    IF ((x0 = FALSE) AND  (x1 = FALSE) AND  (x2 = FALSE) AND  (t0.Q = FALSE)) THEN 
        cstate58 := 7390; y0 := FALSE; y1 := TRUE; t0_start := FALSE; 
    ELSIF ((x0 = FALSE) AND  (x1 = FALSE) AND  (x2 = FALSE) AND  (t0.Q = TRUE)) THEN 
        cstate58 := 7378; y0 := FALSE; y1 := TRUE; t0_start := FALSE; 
    ELSIF ((x0 = FALSE) AND  (x1 = FALSE) AND  (x2 = TRUE) AND  (t0.Q = FALSE)) THEN 
        cstate58 := 7582; y0 := FALSE; y1 := TRUE; t0_start := FALSE; 
    ELSIF ((x0 = FALSE) AND  (x1 = FALSE) AND  (x2 = TRUE) AND  (t0.Q = TRUE)) THEN 
        cstate58 := 7570; y0 := FALSE; y1 := TRUE; t0_start := FALSE; 
    ELSIF ((x0 = FALSE) AND  (x1 = TRUE) AND  (x2 = FALSE) AND  (t0.Q = FALSE)) THEN 
        cstate58 := 6340; y0 := FALSE; y1 := FALSE; t0_start := FALSE; 
    ELSIF ((x0 = FALSE) AND  (x1 = TRUE) AND  (x2 = FALSE) AND  (t0.Q = TRUE)) THEN 
        cstate58 := 6338; y0 := FALSE; y1 := FALSE; t0_start := FALSE; 
    ELSIF ((x0 = FALSE) AND  (x1 = TRUE) AND  (x2 = TRUE) AND  (t0.Q = FALSE)) THEN 
        cstate58 := 6532; y0 := FALSE; y1 := FALSE; t0_start := FALSE; 
    ELSIF ((x0 = FALSE) AND  (x1 = TRUE) AND  (x2 = TRUE) AND  (t0.Q = TRUE)) THEN 
        cstate58 := 6530; y0 := FALSE; y1 := FALSE; t0_start := FALSE; 
    ELSIF ((x0 = TRUE) AND  (x1 = FALSE) AND  (x2 = FALSE) AND  (t0.Q = FALSE)) THEN 
        cstate58 := 5192; y0 := TRUE; y1 := FALSE; t0_start := FALSE; 
    ELSIF ((x0 = TRUE) AND  (x1 = FALSE) AND  (x2 = FALSE) AND  (t0.Q = TRUE)) THEN 
        cstate58 := 5186; y0 := TRUE; y1 := FALSE; t0_start := FALSE; 
    ELSIF ((x0 = TRUE) AND  (x1 = FALSE) AND  (x2 = TRUE) AND  (t0.Q = FALSE)) THEN 
        cstate58 := 3848; y0 := FALSE; y1 := FALSE; t0_start := FALSE; 
    ELSIF ((x0 = TRUE) AND  (x1 = FALSE) AND  (x2 = TRUE) AND  (t0.Q = TRUE)) THEN 
        cstate58 := 3842; y0 := FALSE; y1 := FALSE; t0_start := FALSE; 
    ELSIF ((x0 = TRUE) AND  (x1 = TRUE) AND  (x2 = FALSE) AND  (t0.Q = FALSE)) THEN 
        cstate58 := 4678; y0 := TRUE; y1 := FALSE; t0_start := FALSE; 
    ELSIF ((x0 = TRUE) AND  (x1 = TRUE) AND  (x2 = FALSE) AND  (t0.Q = TRUE)) THEN 
        cstate58 := 4674; y0 := TRUE; y1 := FALSE; t0_start := FALSE; 
    ELSIF ((x0 = TRUE) AND  (x1 = TRUE) AND  (x2 = TRUE) AND  (t0.Q = FALSE)) THEN 
        cstate58 := 2502; y0 := FALSE; y1 := FALSE; t0_start := FALSE; 
    ELSIF ((x0 = TRUE) AND  (x1 = TRUE) AND  (x2 = TRUE) AND  (t0.Q = TRUE)) THEN 
        cstate58 := 2498; y0 := FALSE; y1 := FALSE; t0_start := FALSE; 
    END_IF;
6338:
    IF ((x0 = FALSE) AND  (x1 = FALSE) AND  (x2 = FALSE) AND  (t0.Q = FALSE)) THEN 
        cstate58 := 6340; y0 := FALSE; y1 := FALSE; t0_start := FALSE; 
    ELSIF ((x0 = FALSE) AND  (x1 = FALSE) AND  (x2 = FALSE) AND  (t0.Q = TRUE)) THEN 
        cstate58 := 6338; y0 := FALSE; y1 := FALSE; t0_start := FALSE; 
    ELSIF ((x0 = FALSE) AND  (x1 = FALSE) AND  (x2 = TRUE) AND  (t0.Q = FALSE)) THEN 
        cstate58 := 6468; y0 := FALSE; y1 := FALSE; t0_start := TRUE; t0_up := FALSE; 
    ELSIF ((x0 = FALSE) AND  (x1 = FALSE) AND  (x2 = TRUE) AND  (t0.Q = TRUE)) THEN 
        cstate58 := 6466; y0 := FALSE; y1 := FALSE; t0_start := TRUE; t0_up := FALSE; 
    ELSIF ((x0 = FALSE) AND  (x1 = TRUE) AND  (x2 = FALSE) AND  (t0.Q = FALSE)) THEN 
        cstate58 := 6340; y0 := FALSE; y1 := FALSE; t0_start := FALSE; 
    ELSIF ((x0 = FALSE) AND  (x1 = TRUE) AND  (x2 = FALSE) AND  (t0.Q = TRUE)) THEN 
        cstate58 := 6338; y0 := FALSE; y1 := FALSE; t0_start := FALSE; 
    ELSIF ((x0 = FALSE) AND  (x1 = TRUE) AND  (x2 = TRUE) AND  (t0.Q = FALSE)) THEN 
        cstate58 := 6468; y0 := FALSE; y1 := FALSE; t0_start := TRUE; t0_up := FALSE; 
    ELSIF ((x0 = FALSE) AND  (x1 = TRUE) AND  (x2 = TRUE) AND  (t0.Q = TRUE)) THEN 
        cstate58 := 6466; y0 := FALSE; y1 := FALSE; t0_start := TRUE; t0_up := FALSE; 
    ELSIF ((x0 = TRUE) AND  (x1 = FALSE) AND  (x2 = FALSE) AND  (t0.Q = FALSE)) THEN 
        cstate58 := 4168; y0 := TRUE; y1 := FALSE; t0_start := FALSE; 
    ELSIF ((x0 = TRUE) AND  (x1 = FALSE) AND  (x2 = FALSE) AND  (t0.Q = TRUE)) THEN 
        cstate58 := 4162; y0 := TRUE; y1 := FALSE; t0_start := FALSE; 
    ELSIF ((x0 = TRUE) AND  (x1 = FALSE) AND  (x2 = TRUE) AND  (t0.Q = FALSE)) THEN 
        cstate58 := 2760; y0 := FALSE; y1 := FALSE; t0_start := TRUE; t0_up := FALSE; 
    ELSIF ((x0 = TRUE) AND  (x1 = FALSE) AND  (x2 = TRUE) AND  (t0.Q = TRUE)) THEN 
        cstate58 := 2754; y0 := FALSE; y1 := FALSE; t0_start := TRUE; t0_up := FALSE; 
    ELSIF ((x0 = TRUE) AND  (x1 = TRUE) AND  (x2 = FALSE) AND  (t0.Q = FALSE)) THEN 
        cstate58 := 4678; y0 := TRUE; y1 := FALSE; t0_start := FALSE; 
    ELSIF ((x0 = TRUE) AND  (x1 = TRUE) AND  (x2 = FALSE) AND  (t0.Q = TRUE)) THEN 
        cstate58 := 4674; y0 := TRUE; y1 := FALSE; t0_start := FALSE; 
    ELSIF ((x0 = TRUE) AND  (x1 = TRUE) AND  (x2 = TRUE) AND  (t0.Q = FALSE)) THEN 
        cstate58 := 2566; y0 := FALSE; y1 := FALSE; t0_start := TRUE; t0_up := FALSE; 
    ELSIF ((x0 = TRUE) AND  (x1 = TRUE) AND  (x2 = TRUE) AND  (t0.Q = TRUE)) THEN 
        cstate58 := 2562; y0 := FALSE; y1 := FALSE; t0_start := TRUE; t0_up := FALSE; 
    END_IF;
1226:
    IF ((x0 = FALSE) AND  (x1 = FALSE) AND  (x2 = FALSE) AND  (t0.Q = FALSE)) THEN 
        cstate58 := 1238; y0 := FALSE; y1 := TRUE; t0_start := FALSE; 
    ELSIF ((x0 = FALSE) AND  (x1 = FALSE) AND  (x2 = FALSE) AND  (t0.Q = TRUE)) THEN 
        cstate58 := 1226; y0 := FALSE; y1 := TRUE; t0_start := FALSE; 
    ELSIF ((x0 = FALSE) AND  (x1 = FALSE) AND  (x2 = TRUE) AND  (t0.Q = FALSE)) THEN 
        cstate58 := 1368; y0 := FALSE; y1 := TRUE; t0_start := TRUE; t0_up := FALSE; 
    ELSIF ((x0 = FALSE) AND  (x1 = FALSE) AND  (x2 = TRUE) AND  (t0.Q = TRUE)) THEN 
        cstate58 := 1356; y0 := FALSE; y1 := TRUE; t0_start := TRUE; t0_up := FALSE; 
    ELSIF ((x0 = FALSE) AND  (x1 = TRUE) AND  (x2 = FALSE) AND  (t0.Q = FALSE)) THEN 
        cstate58 := 1220; y0 := FALSE; y1 := FALSE; t0_start := FALSE; 
    ELSIF ((x0 = FALSE) AND  (x1 = TRUE) AND  (x2 = FALSE) AND  (t0.Q = TRUE)) THEN 
        cstate58 := 1218; y0 := FALSE; y1 := FALSE; t0_start := FALSE; 
    ELSIF ((x0 = FALSE) AND  (x1 = TRUE) AND  (x2 = TRUE) AND  (t0.Q = FALSE)) THEN 
        cstate58 := 1348; y0 := FALSE; y1 := FALSE; t0_start := TRUE; t0_up := FALSE; 
    ELSIF ((x0 = FALSE) AND  (x1 = TRUE) AND  (x2 = TRUE) AND  (t0.Q = TRUE)) THEN 
        cstate58 := 1346; y0 := FALSE; y1 := FALSE; t0_start := TRUE; t0_up := FALSE; 
    ELSIF ((x0 = TRUE) AND  (x1 = FALSE) AND  (x2 = FALSE) AND  (t0.Q = FALSE)) THEN 
        cstate58 := 5192; y0 := TRUE; y1 := FALSE; t0_start := FALSE; 
    ELSIF ((x0 = TRUE) AND  (x1 = FALSE) AND  (x2 = FALSE) AND  (t0.Q = TRUE)) THEN 
        cstate58 := 5186; y0 := TRUE; y1 := FALSE; t0_start := FALSE; 
    ELSIF ((x0 = TRUE) AND  (x1 = FALSE) AND  (x2 = TRUE) AND  (t0.Q = FALSE)) THEN 
        cstate58 := 3784; y0 := FALSE; y1 := FALSE; t0_start := TRUE; t0_up := FALSE; 
    ELSIF ((x0 = TRUE) AND  (x1 = FALSE) AND  (x2 = TRUE) AND  (t0.Q = TRUE)) THEN 
        cstate58 := 3778; y0 := FALSE; y1 := FALSE; t0_start := TRUE; t0_up := FALSE; 
    ELSIF ((x0 = TRUE) AND  (x1 = TRUE) AND  (x2 = FALSE) AND  (t0.Q = FALSE)) THEN 
        cstate58 := 4678; y0 := TRUE; y1 := FALSE; t0_start := FALSE; 
    ELSIF ((x0 = TRUE) AND  (x1 = TRUE) AND  (x2 = FALSE) AND  (t0.Q = TRUE)) THEN 
        cstate58 := 4674; y0 := TRUE; y1 := FALSE; t0_start := FALSE; 
    ELSIF ((x0 = TRUE) AND  (x1 = TRUE) AND  (x2 = TRUE) AND  (t0.Q = FALSE)) THEN 
        cstate58 := 2566; y0 := FALSE; y1 := FALSE; t0_start := TRUE; t0_up := FALSE; 
    ELSIF ((x0 = TRUE) AND  (x1 = TRUE) AND  (x2 = TRUE) AND  (t0.Q = TRUE)) THEN 
        cstate58 := 2562; y0 := FALSE; y1 := FALSE; t0_start := TRUE; t0_up := FALSE; 
    END_IF;
7370:
    IF ((x0 = FALSE) AND  (x1 = FALSE) AND  (x2 = FALSE) AND  (t0.Q = FALSE)) THEN 
        cstate58 := 7382; y0 := FALSE; y1 := TRUE; t0_start := FALSE; 
    ELSIF ((x0 = FALSE) AND  (x1 = FALSE) AND  (x2 = FALSE) AND  (t0.Q = TRUE)) THEN 
        cstate58 := 7370; y0 := FALSE; y1 := TRUE; t0_start := FALSE; 
    ELSIF ((x0 = FALSE) AND  (x1 = FALSE) AND  (x2 = TRUE) AND  (t0.Q = FALSE)) THEN 
        cstate58 := 7512; y0 := FALSE; y1 := TRUE; t0_start := TRUE; t0_up := FALSE; 
    ELSIF ((x0 = FALSE) AND  (x1 = FALSE) AND  (x2 = TRUE) AND  (t0.Q = TRUE)) THEN 
        cstate58 := 7500; y0 := FALSE; y1 := TRUE; t0_start := TRUE; t0_up := FALSE; 
    ELSIF ((x0 = FALSE) AND  (x1 = TRUE) AND  (x2 = FALSE) AND  (t0.Q = FALSE)) THEN 
        cstate58 := 6340; y0 := FALSE; y1 := FALSE; t0_start := FALSE; 
    ELSIF ((x0 = FALSE) AND  (x1 = TRUE) AND  (x2 = FALSE) AND  (t0.Q = TRUE)) THEN 
        cstate58 := 6338; y0 := FALSE; y1 := FALSE; t0_start := FALSE; 
    ELSIF ((x0 = FALSE) AND  (x1 = TRUE) AND  (x2 = TRUE) AND  (t0.Q = FALSE)) THEN 
        cstate58 := 6468; y0 := FALSE; y1 := FALSE; t0_start := TRUE; t0_up := FALSE; 
    ELSIF ((x0 = FALSE) AND  (x1 = TRUE) AND  (x2 = TRUE) AND  (t0.Q = TRUE)) THEN 
        cstate58 := 6466; y0 := FALSE; y1 := FALSE; t0_start := TRUE; t0_up := FALSE; 
    ELSIF ((x0 = TRUE) AND  (x1 = FALSE) AND  (x2 = FALSE) AND  (t0.Q = FALSE)) THEN 
        cstate58 := 5192; y0 := TRUE; y1 := FALSE; t0_start := FALSE; 
    ELSIF ((x0 = TRUE) AND  (x1 = FALSE) AND  (x2 = FALSE) AND  (t0.Q = TRUE)) THEN 
        cstate58 := 5186; y0 := TRUE; y1 := FALSE; t0_start := FALSE; 
    ELSIF ((x0 = TRUE) AND  (x1 = FALSE) AND  (x2 = TRUE) AND  (t0.Q = FALSE)) THEN 
        cstate58 := 3784; y0 := FALSE; y1 := FALSE; t0_start := TRUE; t0_up := FALSE; 
    ELSIF ((x0 = TRUE) AND  (x1 = FALSE) AND  (x2 = TRUE) AND  (t0.Q = TRUE)) THEN 
        cstate58 := 3778; y0 := FALSE; y1 := FALSE; t0_start := TRUE; t0_up := FALSE; 
    ELSIF ((x0 = TRUE) AND  (x1 = TRUE) AND  (x2 = FALSE) AND  (t0.Q = FALSE)) THEN 
        cstate58 := 4678; y0 := TRUE; y1 := FALSE; t0_start := FALSE; 
    ELSIF ((x0 = TRUE) AND  (x1 = TRUE) AND  (x2 = FALSE) AND  (t0.Q = TRUE)) THEN 
        cstate58 := 4674; y0 := TRUE; y1 := FALSE; t0_start := FALSE; 
    ELSIF ((x0 = TRUE) AND  (x1 = TRUE) AND  (x2 = TRUE) AND  (t0.Q = FALSE)) THEN 
        cstate58 := 2566; y0 := FALSE; y1 := FALSE; t0_start := TRUE; t0_up := FALSE; 
    ELSIF ((x0 = TRUE) AND  (x1 = TRUE) AND  (x2 = TRUE) AND  (t0.Q = TRUE)) THEN 
        cstate58 := 2562; y0 := FALSE; y1 := FALSE; t0_start := TRUE; t0_up := FALSE; 
    END_IF;
6542:
    IF ((x0 = FALSE) AND  (x1 = FALSE) AND  (x2 = FALSE) AND  (t0.Q = FALSE)) THEN 
        cstate58 := 6362; y0 := FALSE; y1 := TRUE; t0_start := FALSE; 
    ELSIF ((x0 = FALSE) AND  (x1 = FALSE) AND  (x2 = FALSE) AND  (t0.Q = TRUE)) THEN 
        cstate58 := 6350; y0 := FALSE; y1 := TRUE; t0_start := FALSE; 
    ELSIF ((x0 = FALSE) AND  (x1 = FALSE) AND  (x2 = TRUE) AND  (t0.Q = FALSE)) THEN 
        cstate58 := 6554; y0 := FALSE; y1 := TRUE; t0_start := FALSE; 
    ELSIF ((x0 = FALSE) AND  (x1 = FALSE) AND  (x2 = TRUE) AND  (t0.Q = TRUE)) THEN 
        cstate58 := 6542; y0 := FALSE; y1 := TRUE; t0_start := FALSE; 
    ELSIF ((x0 = FALSE) AND  (x1 = TRUE) AND  (x2 = FALSE) AND  (t0.Q = FALSE)) THEN 
        cstate58 := 6340; y0 := FALSE; y1 := FALSE; t0_start := FALSE; 
    ELSIF ((x0 = FALSE) AND  (x1 = TRUE) AND  (x2 = FALSE) AND  (t0.Q = TRUE)) THEN 
        cstate58 := 6338; y0 := FALSE; y1 := FALSE; t0_start := FALSE; 
    ELSIF ((x0 = FALSE) AND  (x1 = TRUE) AND  (x2 = TRUE) AND  (t0.Q = FALSE)) THEN 
        cstate58 := 6532; y0 := FALSE; y1 := FALSE; t0_start := FALSE; 
    ELSIF ((x0 = FALSE) AND  (x1 = TRUE) AND  (x2 = TRUE) AND  (t0.Q = TRUE)) THEN 
        cstate58 := 6530; y0 := FALSE; y1 := FALSE; t0_start := FALSE; 
    ELSIF ((x0 = TRUE) AND  (x1 = FALSE) AND  (x2 = FALSE) AND  (t0.Q = FALSE)) THEN 
        cstate58 := 4168; y0 := TRUE; y1 := FALSE; t0_start := FALSE; 
    ELSIF ((x0 = TRUE) AND  (x1 = FALSE) AND  (x2 = FALSE) AND  (t0.Q = TRUE)) THEN 
        cstate58 := 4162; y0 := TRUE; y1 := FALSE; t0_start := FALSE; 
    ELSIF ((x0 = TRUE) AND  (x1 = FALSE) AND  (x2 = TRUE) AND  (t0.Q = FALSE)) THEN 
        cstate58 := 2824; y0 := FALSE; y1 := FALSE; t0_start := FALSE; 
    ELSIF ((x0 = TRUE) AND  (x1 = FALSE) AND  (x2 = TRUE) AND  (t0.Q = TRUE)) THEN 
        cstate58 := 2818; y0 := FALSE; y1 := FALSE; t0_start := FALSE; 
    ELSIF ((x0 = TRUE) AND  (x1 = TRUE) AND  (x2 = FALSE) AND  (t0.Q = FALSE)) THEN 
        cstate58 := 4678; y0 := TRUE; y1 := FALSE; t0_start := FALSE; 
    ELSIF ((x0 = TRUE) AND  (x1 = TRUE) AND  (x2 = FALSE) AND  (t0.Q = TRUE)) THEN 
        cstate58 := 4674; y0 := TRUE; y1 := FALSE; t0_start := FALSE; 
    ELSIF ((x0 = TRUE) AND  (x1 = TRUE) AND  (x2 = TRUE) AND  (t0.Q = FALSE)) THEN 
        cstate58 := 2502; y0 := FALSE; y1 := FALSE; t0_start := FALSE; 
    ELSIF ((x0 = TRUE) AND  (x1 = TRUE) AND  (x2 = TRUE) AND  (t0.Q = TRUE)) THEN 
        cstate58 := 2498; y0 := FALSE; y1 := FALSE; t0_start := FALSE; 
    END_IF;
4678:
    IF ((x0 = FALSE) AND  ( TRUE ) AND  (x2 = FALSE) AND  (t0.Q = FALSE)) THEN 
        cstate58 := 8388; y0 := TRUE; y1 := FALSE; t0_start := FALSE; 
    ELSIF ((x0 = FALSE) AND  ( TRUE ) AND  (x2 = FALSE) AND  (t0.Q = TRUE)) THEN 
        cstate58 := 8386; y0 := TRUE; y1 := FALSE; t0_start := FALSE; 
    ELSIF ((x0 = FALSE) AND  (x1 = FALSE) AND  (x2 = TRUE) AND  (t0.Q = FALSE)) THEN 
        cstate58 := 6468; y0 := FALSE; y1 := FALSE; t0_start := TRUE; t0_up := FALSE; 
    ELSIF ((x0 = FALSE) AND  (x1 = FALSE) AND  (x2 = TRUE) AND  (t0.Q = TRUE)) THEN 
        cstate58 := 6480; y0 := FALSE; y1 := TRUE; t0_start := TRUE; t0_up := FALSE; 
    ELSIF ((x0 = FALSE) AND  (x1 = TRUE) AND  (x2 = TRUE) AND  (t0.Q = FALSE)) THEN 
        cstate58 := 6468; y0 := FALSE; y1 := FALSE; t0_start := TRUE; t0_up := FALSE; 
    ELSIF ((x0 = FALSE) AND  (x1 = TRUE) AND  (x2 = TRUE) AND  (t0.Q = TRUE)) THEN 
        cstate58 := 6466; y0 := FALSE; y1 := FALSE; t0_start := TRUE; t0_up := FALSE; 
    ELSIF ((x0 = TRUE) AND  (x1 = FALSE) AND  (x2 = FALSE) AND  (t0.Q = FALSE)) THEN 
        cstate58 := 4168; y0 := TRUE; y1 := FALSE; t0_start := FALSE; 
    ELSIF ((x0 = TRUE) AND  (x1 = FALSE) AND  (x2 = FALSE) AND  (t0.Q = TRUE)) THEN 
        cstate58 := 4162; y0 := TRUE; y1 := FALSE; t0_start := FALSE; 
    ELSIF ((x0 = TRUE) AND  (x1 = FALSE) AND  (x2 = TRUE) AND  (t0.Q = FALSE)) THEN 
        cstate58 := 2760; y0 := FALSE; y1 := FALSE; t0_start := TRUE; t0_up := FALSE; 
    ELSIF ((x0 = TRUE) AND  (x1 = FALSE) AND  (x2 = TRUE) AND  (t0.Q = TRUE)) THEN 
        cstate58 := 2754; y0 := FALSE; y1 := FALSE; t0_start := TRUE; t0_up := FALSE; 
    ELSIF ((x0 = TRUE) AND  (x1 = TRUE) AND  (x2 = FALSE) AND  (t0.Q = FALSE)) THEN 
        cstate58 := 4678; y0 := TRUE; y1 := FALSE; t0_start := FALSE; 
    ELSIF ((x0 = TRUE) AND  (x1 = TRUE) AND  (x2 = FALSE) AND  (t0.Q = TRUE)) THEN 
        cstate58 := 4674; y0 := TRUE; y1 := FALSE; t0_start := FALSE; 
    ELSIF ((x0 = TRUE) AND  (x1 = TRUE) AND  (x2 = TRUE) AND  (t0.Q = FALSE)) THEN 
        cstate58 := 2566; y0 := FALSE; y1 := FALSE; t0_start := TRUE; t0_up := FALSE; 
    ELSIF ((x0 = TRUE) AND  (x1 = TRUE) AND  (x2 = TRUE) AND  (t0.Q = TRUE)) THEN 
        cstate58 := 2562; y0 := FALSE; y1 := FALSE; t0_start := TRUE; t0_up := FALSE; 
    END_IF;
9476:
    IF ((x0 = FALSE) AND  (x1 = FALSE) AND  (x2 = FALSE) AND  (t0.Q = FALSE)) THEN 
        cstate58 := 9476; y0 := TRUE; y1 := FALSE; t0_start := FALSE; 
    ELSIF ((x0 = FALSE) AND  (x1 = FALSE) AND  (x2 = FALSE) AND  (t0.Q = TRUE)) THEN 
        cstate58 := 9410; y0 := TRUE; y1 := FALSE; t0_start := FALSE; 
    ELSIF ((x0 = FALSE) AND  (x1 = FALSE) AND  (x2 = TRUE) AND  (t0.Q = FALSE)) THEN 
        cstate58 := 7492; y0 := FALSE; y1 := FALSE; t0_start := TRUE; t0_up := FALSE; 
    ELSIF ((x0 = FALSE) AND  (x1 = FALSE) AND  (x2 = TRUE) AND  (t0.Q = TRUE)) THEN 
        cstate58 := 7500; y0 := FALSE; y1 := TRUE; t0_start := TRUE; t0_up := FALSE; 
    ELSIF ((x0 = FALSE) AND  (x1 = TRUE) AND  (x2 = FALSE) AND  (t0.Q = FALSE)) THEN 
        cstate58 := 8452; y0 := TRUE; y1 := FALSE; t0_start := FALSE; 
    ELSIF ((x0 = FALSE) AND  (x1 = TRUE) AND  (x2 = FALSE) AND  (t0.Q = TRUE)) THEN 
        cstate58 := 8386; y0 := TRUE; y1 := FALSE; t0_start := FALSE; 
    ELSIF ((x0 = FALSE) AND  (x1 = TRUE) AND  (x2 = TRUE) AND  (t0.Q = FALSE)) THEN 
        cstate58 := 6468; y0 := FALSE; y1 := FALSE; t0_start := TRUE; t0_up := FALSE; 
    ELSIF ((x0 = FALSE) AND  (x1 = TRUE) AND  (x2 = TRUE) AND  (t0.Q = TRUE)) THEN 
        cstate58 := 6466; y0 := FALSE; y1 := FALSE; t0_start := TRUE; t0_up := FALSE; 
    ELSIF ((x0 = TRUE) AND  (x1 = FALSE) AND  (x2 = FALSE) AND  (t0.Q = FALSE)) THEN 
        cstate58 := 5256; y0 := TRUE; y1 := FALSE; t0_start := FALSE; 
    ELSIF ((x0 = TRUE) AND  (x1 = FALSE) AND  (x2 = FALSE) AND  (t0.Q = TRUE)) THEN 
        cstate58 := 5186; y0 := TRUE; y1 := FALSE; t0_start := FALSE; 
    ELSIF ((x0 = TRUE) AND  (x1 = FALSE) AND  (x2 = TRUE) AND  (t0.Q = FALSE)) THEN 
        cstate58 := 3784; y0 := FALSE; y1 := FALSE; t0_start := TRUE; t0_up := FALSE; 
    ELSIF ((x0 = TRUE) AND  (x1 = FALSE) AND  (x2 = TRUE) AND  (t0.Q = TRUE)) THEN 
        cstate58 := 3778; y0 := FALSE; y1 := FALSE; t0_start := TRUE; t0_up := FALSE; 
    ELSIF ((x0 = TRUE) AND  (x1 = TRUE) AND  (x2 = FALSE) AND  (t0.Q = FALSE)) THEN 
        cstate58 := 4742; y0 := TRUE; y1 := FALSE; t0_start := FALSE; 
    ELSIF ((x0 = TRUE) AND  (x1 = TRUE) AND  (x2 = FALSE) AND  (t0.Q = TRUE)) THEN 
        cstate58 := 4674; y0 := TRUE; y1 := FALSE; t0_start := FALSE; 
    ELSIF ((x0 = TRUE) AND  (x1 = TRUE) AND  (x2 = TRUE) AND  (t0.Q = FALSE)) THEN 
        cstate58 := 2566; y0 := FALSE; y1 := FALSE; t0_start := TRUE; t0_up := FALSE; 
    ELSIF ((x0 = TRUE) AND  (x1 = TRUE) AND  (x2 = TRUE) AND  (t0.Q = TRUE)) THEN 
        cstate58 := 2562; y0 := FALSE; y1 := FALSE; t0_start := TRUE; t0_up := FALSE; 
    END_IF;
7378:
    IF ((x0 = FALSE) AND  (x1 = FALSE) AND  (x2 = FALSE) AND  (t0.Q = FALSE)) THEN 
        cstate58 := 7390; y0 := FALSE; y1 := TRUE; t0_start := FALSE; 
    ELSIF ((x0 = FALSE) AND  (x1 = FALSE) AND  (x2 = FALSE) AND  (t0.Q = TRUE)) THEN 
        cstate58 := 7378; y0 := FALSE; y1 := TRUE; t0_start := FALSE; 
    ELSIF ((x0 = FALSE) AND  (x1 = FALSE) AND  (x2 = TRUE) AND  (t0.Q = FALSE)) THEN 
        cstate58 := 7520; y0 := FALSE; y1 := TRUE; t0_start := TRUE; t0_up := FALSE; 
    ELSIF ((x0 = FALSE) AND  (x1 = FALSE) AND  (x2 = TRUE) AND  (t0.Q = TRUE)) THEN 
        cstate58 := 7508; y0 := FALSE; y1 := TRUE; t0_start := TRUE; t0_up := FALSE; 
    ELSIF ((x0 = FALSE) AND  (x1 = TRUE) AND  (x2 = FALSE) AND  (t0.Q = FALSE)) THEN 
        cstate58 := 6340; y0 := FALSE; y1 := FALSE; t0_start := FALSE; 
    ELSIF ((x0 = FALSE) AND  (x1 = TRUE) AND  (x2 = FALSE) AND  (t0.Q = TRUE)) THEN 
        cstate58 := 6338; y0 := FALSE; y1 := FALSE; t0_start := FALSE; 
    ELSIF ((x0 = FALSE) AND  (x1 = TRUE) AND  (x2 = TRUE) AND  (t0.Q = FALSE)) THEN 
        cstate58 := 6468; y0 := FALSE; y1 := FALSE; t0_start := TRUE; t0_up := FALSE; 
    ELSIF ((x0 = FALSE) AND  (x1 = TRUE) AND  (x2 = TRUE) AND  (t0.Q = TRUE)) THEN 
        cstate58 := 6466; y0 := FALSE; y1 := FALSE; t0_start := TRUE; t0_up := FALSE; 
    ELSIF ((x0 = TRUE) AND  (x1 = FALSE) AND  (x2 = FALSE) AND  (t0.Q = FALSE)) THEN 
        cstate58 := 5192; y0 := TRUE; y1 := FALSE; t0_start := FALSE; 
    ELSIF ((x0 = TRUE) AND  (x1 = FALSE) AND  (x2 = FALSE) AND  (t0.Q = TRUE)) THEN 
        cstate58 := 5186; y0 := TRUE; y1 := FALSE; t0_start := FALSE; 
    ELSIF ((x0 = TRUE) AND  (x1 = FALSE) AND  (x2 = TRUE) AND  (t0.Q = FALSE)) THEN 
        cstate58 := 3784; y0 := FALSE; y1 := FALSE; t0_start := TRUE; t0_up := FALSE; 
    ELSIF ((x0 = TRUE) AND  (x1 = FALSE) AND  (x2 = TRUE) AND  (t0.Q = TRUE)) THEN 
        cstate58 := 3778; y0 := FALSE; y1 := FALSE; t0_start := TRUE; t0_up := FALSE; 
    ELSIF ((x0 = TRUE) AND  (x1 = TRUE) AND  (x2 = FALSE) AND  (t0.Q = FALSE)) THEN 
        cstate58 := 4678; y0 := TRUE; y1 := FALSE; t0_start := FALSE; 
    ELSIF ((x0 = TRUE) AND  (x1 = TRUE) AND  (x2 = FALSE) AND  (t0.Q = TRUE)) THEN 
        cstate58 := 4674; y0 := TRUE; y1 := FALSE; t0_start := FALSE; 
    ELSIF ((x0 = TRUE) AND  (x1 = TRUE) AND  (x2 = TRUE) AND  (t0.Q = FALSE)) THEN 
        cstate58 := 2566; y0 := FALSE; y1 := FALSE; t0_start := TRUE; t0_up := FALSE; 
    ELSIF ((x0 = TRUE) AND  (x1 = TRUE) AND  (x2 = TRUE) AND  (t0.Q = TRUE)) THEN 
        cstate58 := 2562; y0 := FALSE; y1 := FALSE; t0_start := TRUE; t0_up := FALSE; 
    END_IF;
1368:
    IF ((x0 = FALSE) AND  (x1 = FALSE) AND  (x2 = FALSE) AND  (t0.Q = FALSE)) THEN 
        cstate58 := 1304; y0 := FALSE; y1 := TRUE; t0_start := FALSE; 
    ELSIF ((x0 = FALSE) AND  (x1 = FALSE) AND  (x2 = FALSE) AND  (t0.Q = TRUE)) THEN 
        cstate58 := 1226; y0 := FALSE; y1 := TRUE; t0_start := FALSE; 
    ELSIF ((x0 = FALSE) AND  (x1 = FALSE) AND  (x2 = TRUE) AND  (t0.Q = FALSE)) THEN 
        cstate58 := 1368; y0 := FALSE; y1 := TRUE; t0_start := FALSE; 
    ELSIF ((x0 = FALSE) AND  (x1 = FALSE) AND  (x2 = TRUE) AND  (t0.Q = TRUE)) THEN 
        cstate58 := 1418; y0 := FALSE; y1 := TRUE; t0_start := FALSE; 
    ELSIF ((x0 = FALSE) AND  (x1 = TRUE) AND  (x2 = FALSE) AND  (t0.Q = FALSE)) THEN 
        cstate58 := 1284; y0 := FALSE; y1 := FALSE; t0_start := FALSE; 
    ELSIF ((x0 = FALSE) AND  (x1 = TRUE) AND  (x2 = FALSE) AND  (t0.Q = TRUE)) THEN 
        cstate58 := 1218; y0 := FALSE; y1 := FALSE; t0_start := FALSE; 
    ELSIF ((x0 = FALSE) AND  (x1 = TRUE) AND  (x2 = TRUE) AND  (t0.Q = FALSE)) THEN 
        cstate58 := 1348; y0 := FALSE; y1 := FALSE; t0_start := FALSE; 
    ELSIF ((x0 = FALSE) AND  (x1 = TRUE) AND  (x2 = TRUE) AND  (t0.Q = TRUE)) THEN 
        cstate58 := 1410; y0 := FALSE; y1 := FALSE; t0_start := FALSE; 
    ELSIF ((x0 = TRUE) AND  (x1 = FALSE) AND  (x2 = FALSE) AND  (t0.Q = FALSE)) THEN 
        cstate58 := 5256; y0 := TRUE; y1 := FALSE; t0_start := FALSE; 
    ELSIF ((x0 = TRUE) AND  (x1 = FALSE) AND  (x2 = FALSE) AND  (t0.Q = TRUE)) THEN 
        cstate58 := 5186; y0 := TRUE; y1 := FALSE; t0_start := FALSE; 
    ELSIF ((x0 = TRUE) AND  (x1 = FALSE) AND  (x2 = TRUE) AND  (t0.Q = FALSE)) THEN 
        cstate58 := 3784; y0 := FALSE; y1 := FALSE; t0_start := FALSE; 
    ELSIF ((x0 = TRUE) AND  (x1 = FALSE) AND  (x2 = TRUE) AND  (t0.Q = TRUE)) THEN 
        cstate58 := 3842; y0 := FALSE; y1 := FALSE; t0_start := FALSE; 
    ELSIF ((x0 = TRUE) AND  (x1 = TRUE) AND  (x2 = FALSE) AND  (t0.Q = FALSE)) THEN 
        cstate58 := 4742; y0 := TRUE; y1 := FALSE; t0_start := FALSE; 
    ELSIF ((x0 = TRUE) AND  (x1 = TRUE) AND  (x2 = FALSE) AND  (t0.Q = TRUE)) THEN 
        cstate58 := 4674; y0 := TRUE; y1 := FALSE; t0_start := FALSE; 
    ELSIF ((x0 = TRUE) AND  (x1 = TRUE) AND  (x2 = TRUE) AND  (t0.Q = FALSE)) THEN 
        cstate58 := 2566; y0 := FALSE; y1 := FALSE; t0_start := FALSE; 
    ELSIF ((x0 = TRUE) AND  (x1 = TRUE) AND  (x2 = TRUE) AND  (t0.Q = TRUE)) THEN 
        cstate58 := 2498; y0 := FALSE; y1 := FALSE; t0_start := FALSE; 
    END_IF;
7562:
    IF ((x0 = FALSE) AND  (x1 = FALSE) AND  (x2 = FALSE) AND  (t0.Q = FALSE)) THEN 
        cstate58 := 7382; y0 := FALSE; y1 := TRUE; t0_start := FALSE; 
    ELSIF ((x0 = FALSE) AND  (x1 = FALSE) AND  (x2 = FALSE) AND  (t0.Q = TRUE)) THEN 
        cstate58 := 7370; y0 := FALSE; y1 := TRUE; t0_start := FALSE; 
    ELSIF ((x0 = FALSE) AND  (x1 = FALSE) AND  (x2 = TRUE) AND  (t0.Q = FALSE)) THEN 
        cstate58 := 7574; y0 := FALSE; y1 := TRUE; t0_start := FALSE; 
    ELSIF ((x0 = FALSE) AND  (x1 = FALSE) AND  (x2 = TRUE) AND  (t0.Q = TRUE)) THEN 
        cstate58 := 7562; y0 := FALSE; y1 := TRUE; t0_start := FALSE; 
    ELSIF ((x0 = FALSE) AND  (x1 = TRUE) AND  (x2 = FALSE) AND  (t0.Q = FALSE)) THEN 
        cstate58 := 6340; y0 := FALSE; y1 := FALSE; t0_start := FALSE; 
    ELSIF ((x0 = FALSE) AND  (x1 = TRUE) AND  (x2 = FALSE) AND  (t0.Q = TRUE)) THEN 
        cstate58 := 6338; y0 := FALSE; y1 := FALSE; t0_start := FALSE; 
    ELSIF ((x0 = FALSE) AND  (x1 = TRUE) AND  (x2 = TRUE) AND  (t0.Q = FALSE)) THEN 
        cstate58 := 6532; y0 := FALSE; y1 := FALSE; t0_start := FALSE; 
    ELSIF ((x0 = FALSE) AND  (x1 = TRUE) AND  (x2 = TRUE) AND  (t0.Q = TRUE)) THEN 
        cstate58 := 6530; y0 := FALSE; y1 := FALSE; t0_start := FALSE; 
    ELSIF ((x0 = TRUE) AND  (x1 = FALSE) AND  (x2 = FALSE) AND  (t0.Q = FALSE)) THEN 
        cstate58 := 5192; y0 := TRUE; y1 := FALSE; t0_start := FALSE; 
    ELSIF ((x0 = TRUE) AND  (x1 = FALSE) AND  (x2 = FALSE) AND  (t0.Q = TRUE)) THEN 
        cstate58 := 5186; y0 := TRUE; y1 := FALSE; t0_start := FALSE; 
    ELSIF ((x0 = TRUE) AND  (x1 = FALSE) AND  (x2 = TRUE) AND  (t0.Q = FALSE)) THEN 
        cstate58 := 3848; y0 := FALSE; y1 := FALSE; t0_start := FALSE; 
    ELSIF ((x0 = TRUE) AND  (x1 = FALSE) AND  (x2 = TRUE) AND  (t0.Q = TRUE)) THEN 
        cstate58 := 3842; y0 := FALSE; y1 := FALSE; t0_start := FALSE; 
    ELSIF ((x0 = TRUE) AND  (x1 = TRUE) AND  (x2 = FALSE) AND  (t0.Q = FALSE)) THEN 
        cstate58 := 4678; y0 := TRUE; y1 := FALSE; t0_start := FALSE; 
    ELSIF ((x0 = TRUE) AND  (x1 = TRUE) AND  (x2 = FALSE) AND  (t0.Q = TRUE)) THEN 
        cstate58 := 4674; y0 := TRUE; y1 := FALSE; t0_start := FALSE; 
    ELSIF ((x0 = TRUE) AND  (x1 = TRUE) AND  (x2 = TRUE) AND  (t0.Q = FALSE)) THEN 
        cstate58 := 2502; y0 := FALSE; y1 := FALSE; t0_start := FALSE; 
    ELSIF ((x0 = TRUE) AND  (x1 = TRUE) AND  (x2 = TRUE) AND  (t0.Q = TRUE)) THEN 
        cstate58 := 2498; y0 := FALSE; y1 := FALSE; t0_start := FALSE; 
    END_IF;
6432:
    IF ((x0 = FALSE) AND  (x1 = FALSE) AND  (x2 = FALSE) AND  (t0.Q = FALSE)) THEN 
        cstate58 := 6432; y0 := FALSE; y1 := TRUE; t0_start := FALSE; 
    ELSIF ((x0 = FALSE) AND  (x1 = FALSE) AND  (x2 = FALSE) AND  (t0.Q = TRUE)) THEN 
        cstate58 := 6354; y0 := FALSE; y1 := TRUE; t0_start := FALSE; 
    ELSIF ((x0 = FALSE) AND  (x1 = FALSE) AND  (x2 = TRUE) AND  (t0.Q = FALSE)) THEN 
        cstate58 := 6496; y0 := FALSE; y1 := TRUE; t0_start := TRUE; t0_up := FALSE; 
    ELSIF ((x0 = FALSE) AND  (x1 = FALSE) AND  (x2 = TRUE) AND  (t0.Q = TRUE)) THEN 
        cstate58 := 6484; y0 := FALSE; y1 := TRUE; t0_start := TRUE; t0_up := FALSE; 
    ELSIF ((x0 = FALSE) AND  (x1 = TRUE) AND  (x2 = FALSE) AND  (t0.Q = FALSE)) THEN 
        cstate58 := 6404; y0 := FALSE; y1 := FALSE; t0_start := FALSE; 
    ELSIF ((x0 = FALSE) AND  (x1 = TRUE) AND  (x2 = FALSE) AND  (t0.Q = TRUE)) THEN 
        cstate58 := 6338; y0 := FALSE; y1 := FALSE; t0_start := FALSE; 
    ELSIF ((x0 = FALSE) AND  (x1 = TRUE) AND  (x2 = TRUE) AND  (t0.Q = FALSE)) THEN 
        cstate58 := 6468; y0 := FALSE; y1 := FALSE; t0_start := TRUE; t0_up := FALSE; 
    ELSIF ((x0 = FALSE) AND  (x1 = TRUE) AND  (x2 = TRUE) AND  (t0.Q = TRUE)) THEN 
        cstate58 := 6466; y0 := FALSE; y1 := FALSE; t0_start := TRUE; t0_up := FALSE; 
    ELSIF ((x0 = TRUE) AND  (x1 = FALSE) AND  (x2 = FALSE) AND  (t0.Q = FALSE)) THEN 
        cstate58 := 4232; y0 := TRUE; y1 := FALSE; t0_start := FALSE; 
    ELSIF ((x0 = TRUE) AND  (x1 = FALSE) AND  (x2 = FALSE) AND  (t0.Q = TRUE)) THEN 
        cstate58 := 4162; y0 := TRUE; y1 := FALSE; t0_start := FALSE; 
    ELSIF ((x0 = TRUE) AND  (x1 = FALSE) AND  (x2 = TRUE) AND  (t0.Q = FALSE)) THEN 
        cstate58 := 2760; y0 := FALSE; y1 := FALSE; t0_start := TRUE; t0_up := FALSE; 
    ELSIF ((x0 = TRUE) AND  (x1 = FALSE) AND  (x2 = TRUE) AND  (t0.Q = TRUE)) THEN 
        cstate58 := 2754; y0 := FALSE; y1 := FALSE; t0_start := TRUE; t0_up := FALSE; 
    ELSIF ((x0 = TRUE) AND  (x1 = TRUE) AND  (x2 = FALSE) AND  (t0.Q = FALSE)) THEN 
        cstate58 := 4742; y0 := TRUE; y1 := FALSE; t0_start := FALSE; 
    ELSIF ((x0 = TRUE) AND  (x1 = TRUE) AND  (x2 = FALSE) AND  (t0.Q = TRUE)) THEN 
        cstate58 := 4674; y0 := TRUE; y1 := FALSE; t0_start := FALSE; 
    ELSIF ((x0 = TRUE) AND  (x1 = TRUE) AND  (x2 = TRUE) AND  (t0.Q = FALSE)) THEN 
        cstate58 := 2566; y0 := FALSE; y1 := FALSE; t0_start := TRUE; t0_up := FALSE; 
    ELSIF ((x0 = TRUE) AND  (x1 = TRUE) AND  (x2 = TRUE) AND  (t0.Q = TRUE)) THEN 
        cstate58 := 2562; y0 := FALSE; y1 := FALSE; t0_start := TRUE; t0_up := FALSE; 
    END_IF;
5192:
    IF ((x0 = FALSE) AND  (x1 = FALSE) AND  (x2 = FALSE) AND  (t0.Q = FALSE)) THEN 
        cstate58 := 9412; y0 := TRUE; y1 := FALSE; t0_start := FALSE; 
    ELSIF ((x0 = FALSE) AND  (x1 = FALSE) AND  (x2 = FALSE) AND  (t0.Q = TRUE)) THEN 
        cstate58 := 9410; y0 := TRUE; y1 := FALSE; t0_start := FALSE; 
    ELSIF ((x0 = FALSE) AND  (x1 = FALSE) AND  (x2 = TRUE) AND  (t0.Q = FALSE)) THEN 
        cstate58 := 7492; y0 := FALSE; y1 := FALSE; t0_start := TRUE; t0_up := FALSE; 
    ELSIF ((x0 = FALSE) AND  (x1 = FALSE) AND  (x2 = TRUE) AND  (t0.Q = TRUE)) THEN 
        cstate58 := 7508; y0 := FALSE; y1 := TRUE; t0_start := TRUE; t0_up := FALSE; 
    ELSIF ((x0 = FALSE) AND  (x1 = TRUE) AND  (x2 = FALSE) AND  (t0.Q = FALSE)) THEN 
        cstate58 := 8388; y0 := TRUE; y1 := FALSE; t0_start := FALSE; 
    ELSIF ((x0 = FALSE) AND  (x1 = TRUE) AND  (x2 = FALSE) AND  (t0.Q = TRUE)) THEN 
        cstate58 := 8386; y0 := TRUE; y1 := FALSE; t0_start := FALSE; 
    ELSIF ((x0 = FALSE) AND  (x1 = TRUE) AND  (x2 = TRUE) AND  (t0.Q = FALSE)) THEN 
        cstate58 := 6468; y0 := FALSE; y1 := FALSE; t0_start := TRUE; t0_up := FALSE; 
    ELSIF ((x0 = FALSE) AND  (x1 = TRUE) AND  (x2 = TRUE) AND  (t0.Q = TRUE)) THEN 
        cstate58 := 6466; y0 := FALSE; y1 := FALSE; t0_start := TRUE; t0_up := FALSE; 
    ELSIF ((x0 = TRUE) AND  (x1 = FALSE) AND  (x2 = FALSE) AND  (t0.Q = FALSE)) THEN 
        cstate58 := 5192; y0 := TRUE; y1 := FALSE; t0_start := FALSE; 
    ELSIF ((x0 = TRUE) AND  (x1 = FALSE) AND  (x2 = FALSE) AND  (t0.Q = TRUE)) THEN 
        cstate58 := 5186; y0 := TRUE; y1 := FALSE; t0_start := FALSE; 
    ELSIF ((x0 = TRUE) AND  (x1 = FALSE) AND  (x2 = TRUE) AND  (t0.Q = FALSE)) THEN 
        cstate58 := 3784; y0 := FALSE; y1 := FALSE; t0_start := TRUE; t0_up := FALSE; 
    ELSIF ((x0 = TRUE) AND  (x1 = FALSE) AND  (x2 = TRUE) AND  (t0.Q = TRUE)) THEN 
        cstate58 := 3778; y0 := FALSE; y1 := FALSE; t0_start := TRUE; t0_up := FALSE; 
    ELSIF ((x0 = TRUE) AND  (x1 = TRUE) AND  (x2 = FALSE) AND  (t0.Q = FALSE)) THEN 
        cstate58 := 4678; y0 := TRUE; y1 := FALSE; t0_start := FALSE; 
    ELSIF ((x0 = TRUE) AND  (x1 = TRUE) AND  (x2 = FALSE) AND  (t0.Q = TRUE)) THEN 
        cstate58 := 4674; y0 := TRUE; y1 := FALSE; t0_start := FALSE; 
    ELSIF ((x0 = TRUE) AND  (x1 = TRUE) AND  (x2 = TRUE) AND  (t0.Q = FALSE)) THEN 
        cstate58 := 2566; y0 := FALSE; y1 := FALSE; t0_start := TRUE; t0_up := FALSE; 
    ELSIF ((x0 = TRUE) AND  (x1 = TRUE) AND  (x2 = TRUE) AND  (t0.Q = TRUE)) THEN 
        cstate58 := 2562; y0 := FALSE; y1 := FALSE; t0_start := TRUE; t0_up := FALSE; 
    END_IF;
4674:
    IF ((x0 = FALSE) AND  ( TRUE ) AND  (x2 = FALSE) AND  (t0.Q = FALSE)) THEN 
        cstate58 := 8388; y0 := TRUE; y1 := FALSE; t0_start := FALSE; 
    ELSIF ((x0 = FALSE) AND  ( TRUE ) AND  (x2 = FALSE) AND  (t0.Q = TRUE)) THEN 
        cstate58 := 8386; y0 := TRUE; y1 := FALSE; t0_start := FALSE; 
    ELSIF ((x0 = FALSE) AND  (x1 = FALSE) AND  (x2 = TRUE) AND  (t0.Q = FALSE)) THEN 
        cstate58 := 6468; y0 := FALSE; y1 := FALSE; t0_start := TRUE; t0_up := FALSE; 
    ELSIF ((x0 = FALSE) AND  (x1 = FALSE) AND  (x2 = TRUE) AND  (t0.Q = TRUE)) THEN 
        cstate58 := 6466; y0 := FALSE; y1 := FALSE; t0_start := TRUE; t0_up := FALSE; 
    ELSIF ((x0 = FALSE) AND  (x1 = TRUE) AND  (x2 = TRUE) AND  (t0.Q = FALSE)) THEN 
        cstate58 := 6468; y0 := FALSE; y1 := FALSE; t0_start := TRUE; t0_up := FALSE; 
    ELSIF ((x0 = FALSE) AND  (x1 = TRUE) AND  (x2 = TRUE) AND  (t0.Q = TRUE)) THEN 
        cstate58 := 6466; y0 := FALSE; y1 := FALSE; t0_start := TRUE; t0_up := FALSE; 
    ELSIF ((x0 = TRUE) AND  (x1 = FALSE) AND  (x2 = FALSE) AND  (t0.Q = FALSE)) THEN 
        cstate58 := 4168; y0 := TRUE; y1 := FALSE; t0_start := FALSE; 
    ELSIF ((x0 = TRUE) AND  (x1 = FALSE) AND  (x2 = FALSE) AND  (t0.Q = TRUE)) THEN 
        cstate58 := 4162; y0 := TRUE; y1 := FALSE; t0_start := FALSE; 
    ELSIF ((x0 = TRUE) AND  (x1 = FALSE) AND  (x2 = TRUE) AND  (t0.Q = FALSE)) THEN 
        cstate58 := 2760; y0 := FALSE; y1 := FALSE; t0_start := TRUE; t0_up := FALSE; 
    ELSIF ((x0 = TRUE) AND  (x1 = FALSE) AND  (x2 = TRUE) AND  (t0.Q = TRUE)) THEN 
        cstate58 := 2754; y0 := FALSE; y1 := FALSE; t0_start := TRUE; t0_up := FALSE; 
    ELSIF ((x0 = TRUE) AND  (x1 = TRUE) AND  (x2 = FALSE) AND  (t0.Q = FALSE)) THEN 
        cstate58 := 4678; y0 := TRUE; y1 := FALSE; t0_start := FALSE; 
    ELSIF ((x0 = TRUE) AND  (x1 = TRUE) AND  (x2 = FALSE) AND  (t0.Q = TRUE)) THEN 
        cstate58 := 4674; y0 := TRUE; y1 := FALSE; t0_start := FALSE; 
    ELSIF ((x0 = TRUE) AND  (x1 = TRUE) AND  (x2 = TRUE) AND  (t0.Q = FALSE)) THEN 
        cstate58 := 2566; y0 := FALSE; y1 := FALSE; t0_start := TRUE; t0_up := FALSE; 
    ELSIF ((x0 = TRUE) AND  (x1 = TRUE) AND  (x2 = TRUE) AND  (t0.Q = TRUE)) THEN 
        cstate58 := 2562; y0 := FALSE; y1 := FALSE; t0_start := TRUE; t0_up := FALSE; 
    END_IF;
1220:
    IF ((x0 = FALSE) AND  (x1 = FALSE) AND  (x2 = FALSE) AND  (t0.Q = FALSE)) THEN 
        cstate58 := 1220; y0 := FALSE; y1 := FALSE; t0_start := FALSE; 
    ELSIF ((x0 = FALSE) AND  (x1 = FALSE) AND  (x2 = FALSE) AND  (t0.Q = TRUE)) THEN 
        cstate58 := 1226; y0 := FALSE; y1 := TRUE; t0_start := FALSE; 
    ELSIF ((x0 = FALSE) AND  (x1 = FALSE) AND  (x2 = TRUE) AND  (t0.Q = FALSE)) THEN 
        cstate58 := 1348; y0 := FALSE; y1 := FALSE; t0_start := TRUE; t0_up := FALSE; 
    ELSIF ((x0 = FALSE) AND  (x1 = FALSE) AND  (x2 = TRUE) AND  (t0.Q = TRUE)) THEN 
        cstate58 := 1356; y0 := FALSE; y1 := TRUE; t0_start := TRUE; t0_up := FALSE; 
    ELSIF ((x0 = FALSE) AND  (x1 = TRUE) AND  (x2 = FALSE) AND  (t0.Q = FALSE)) THEN 
        cstate58 := 1220; y0 := FALSE; y1 := FALSE; t0_start := FALSE; 
    ELSIF ((x0 = FALSE) AND  (x1 = TRUE) AND  (x2 = FALSE) AND  (t0.Q = TRUE)) THEN 
        cstate58 := 1218; y0 := FALSE; y1 := FALSE; t0_start := FALSE; 
    ELSIF ((x0 = FALSE) AND  (x1 = TRUE) AND  (x2 = TRUE) AND  (t0.Q = FALSE)) THEN 
        cstate58 := 1348; y0 := FALSE; y1 := FALSE; t0_start := TRUE; t0_up := FALSE; 
    ELSIF ((x0 = FALSE) AND  (x1 = TRUE) AND  (x2 = TRUE) AND  (t0.Q = TRUE)) THEN 
        cstate58 := 1346; y0 := FALSE; y1 := FALSE; t0_start := TRUE; t0_up := FALSE; 
    ELSIF ((x0 = TRUE) AND  (x1 = FALSE) AND  (x2 = FALSE) AND  (t0.Q = FALSE)) THEN 
        cstate58 := 5192; y0 := TRUE; y1 := FALSE; t0_start := FALSE; 
    ELSIF ((x0 = TRUE) AND  (x1 = FALSE) AND  (x2 = FALSE) AND  (t0.Q = TRUE)) THEN 
        cstate58 := 5186; y0 := TRUE; y1 := FALSE; t0_start := FALSE; 
    ELSIF ((x0 = TRUE) AND  (x1 = FALSE) AND  (x2 = TRUE) AND  (t0.Q = FALSE)) THEN 
        cstate58 := 3784; y0 := FALSE; y1 := FALSE; t0_start := TRUE; t0_up := FALSE; 
    ELSIF ((x0 = TRUE) AND  (x1 = FALSE) AND  (x2 = TRUE) AND  (t0.Q = TRUE)) THEN 
        cstate58 := 3778; y0 := FALSE; y1 := FALSE; t0_start := TRUE; t0_up := FALSE; 
    ELSIF ((x0 = TRUE) AND  (x1 = TRUE) AND  (x2 = FALSE) AND  (t0.Q = FALSE)) THEN 
        cstate58 := 4678; y0 := TRUE; y1 := FALSE; t0_start := FALSE; 
    ELSIF ((x0 = TRUE) AND  (x1 = TRUE) AND  (x2 = FALSE) AND  (t0.Q = TRUE)) THEN 
        cstate58 := 4674; y0 := TRUE; y1 := FALSE; t0_start := FALSE; 
    ELSIF ((x0 = TRUE) AND  (x1 = TRUE) AND  (x2 = TRUE) AND  (t0.Q = FALSE)) THEN 
        cstate58 := 2566; y0 := FALSE; y1 := FALSE; t0_start := TRUE; t0_up := FALSE; 
    ELSIF ((x0 = TRUE) AND  (x1 = TRUE) AND  (x2 = TRUE) AND  (t0.Q = TRUE)) THEN 
        cstate58 := 2562; y0 := FALSE; y1 := FALSE; t0_start := TRUE; t0_up := FALSE; 
    END_IF;
2694:
    IF ((x0 = FALSE) AND  (x1 = FALSE) AND  (x2 = FALSE) AND  (t0.Q = FALSE)) THEN 
        cstate58 := 6404; y0 := FALSE; y1 := FALSE; t0_start := FALSE; 
    ELSIF ((x0 = FALSE) AND  (x1 = FALSE) AND  (x2 = FALSE) AND  (t0.Q = TRUE)) THEN 
        cstate58 := 6350; y0 := FALSE; y1 := TRUE; t0_start := FALSE; 
    ELSIF ((x0 = FALSE) AND  (x1 = FALSE) AND  (x2 = TRUE) AND  (t0.Q = FALSE)) THEN 
        cstate58 := 6468; y0 := FALSE; y1 := FALSE; t0_start := TRUE; t0_up := FALSE; 
    ELSIF ((x0 = FALSE) AND  (x1 = FALSE) AND  (x2 = TRUE) AND  (t0.Q = TRUE)) THEN 
        cstate58 := 6480; y0 := FALSE; y1 := TRUE; t0_start := TRUE; t0_up := FALSE; 
    ELSIF ((x0 = FALSE) AND  (x1 = TRUE) AND  (x2 = FALSE) AND  (t0.Q = FALSE)) THEN 
        cstate58 := 6404; y0 := FALSE; y1 := FALSE; t0_start := FALSE; 
    ELSIF ((x0 = FALSE) AND  (x1 = TRUE) AND  (x2 = FALSE) AND  (t0.Q = TRUE)) THEN 
        cstate58 := 6338; y0 := FALSE; y1 := FALSE; t0_start := FALSE; 
    ELSIF ((x0 = FALSE) AND  (x1 = TRUE) AND  (x2 = TRUE) AND  (t0.Q = FALSE)) THEN 
        cstate58 := 6468; y0 := FALSE; y1 := FALSE; t0_start := TRUE; t0_up := FALSE; 
    ELSIF ((x0 = FALSE) AND  (x1 = TRUE) AND  (x2 = TRUE) AND  (t0.Q = TRUE)) THEN 
        cstate58 := 6466; y0 := FALSE; y1 := FALSE; t0_start := TRUE; t0_up := FALSE; 
    ELSIF ((x0 = TRUE) AND  (x1 = FALSE) AND  (x2 = FALSE) AND  (t0.Q = FALSE)) THEN 
        cstate58 := 2184; y0 := FALSE; y1 := FALSE; t0_start := FALSE; 
    ELSIF ((x0 = TRUE) AND  (x1 = FALSE) AND  (x2 = FALSE) AND  (t0.Q = TRUE)) THEN 
        cstate58 := 2114; y0 := FALSE; y1 := FALSE; t0_start := FALSE; 
    ELSIF ((x0 = TRUE) AND  (x1 = FALSE) AND  (x2 = TRUE) AND  (t0.Q = FALSE)) THEN 
        cstate58 := 2760; y0 := FALSE; y1 := FALSE; t0_start := TRUE; t0_up := FALSE; 
    ELSIF ((x0 = TRUE) AND  (x1 = FALSE) AND  (x2 = TRUE) AND  (t0.Q = TRUE)) THEN 
        cstate58 := 2754; y0 := FALSE; y1 := FALSE; t0_start := TRUE; t0_up := FALSE; 
    ELSIF ((x0 = TRUE) AND  (x1 = TRUE) AND  (x2 = FALSE) AND  (t0.Q = FALSE)) THEN 
        cstate58 := 2694; y0 := FALSE; y1 := FALSE; t0_start := FALSE; 
    ELSIF ((x0 = TRUE) AND  (x1 = TRUE) AND  (x2 = FALSE) AND  (t0.Q = TRUE)) THEN 
        cstate58 := 2626; y0 := FALSE; y1 := FALSE; t0_start := FALSE; 
    ELSIF ((x0 = TRUE) AND  (x1 = TRUE) AND  (x2 = TRUE) AND  (t0.Q = FALSE)) THEN 
        cstate58 := 2566; y0 := FALSE; y1 := FALSE; t0_start := TRUE; t0_up := FALSE; 
    ELSIF ((x0 = TRUE) AND  (x1 = TRUE) AND  (x2 = TRUE) AND  (t0.Q = TRUE)) THEN 
        cstate58 := 2562; y0 := FALSE; y1 := FALSE; t0_start := TRUE; t0_up := FALSE; 
    END_IF;
6530:
    IF ((x0 = FALSE) AND  (x1 = FALSE) AND  (x2 = FALSE) AND  (t0.Q = FALSE)) THEN 
        cstate58 := 6340; y0 := FALSE; y1 := FALSE; t0_start := FALSE; 
    ELSIF ((x0 = FALSE) AND  (x1 = FALSE) AND  (x2 = FALSE) AND  (t0.Q = TRUE)) THEN 
        cstate58 := 6338; y0 := FALSE; y1 := FALSE; t0_start := FALSE; 
    ELSIF ((x0 = FALSE) AND  (x1 = FALSE) AND  (x2 = TRUE) AND  (t0.Q = FALSE)) THEN 
        cstate58 := 6532; y0 := FALSE; y1 := FALSE; t0_start := FALSE; 
    ELSIF ((x0 = FALSE) AND  (x1 = FALSE) AND  (x2 = TRUE) AND  (t0.Q = TRUE)) THEN 
        cstate58 := 6530; y0 := FALSE; y1 := FALSE; t0_start := FALSE; 
    ELSIF ((x0 = FALSE) AND  (x1 = TRUE) AND  (x2 = FALSE) AND  (t0.Q = FALSE)) THEN 
        cstate58 := 6340; y0 := FALSE; y1 := FALSE; t0_start := FALSE; 
    ELSIF ((x0 = FALSE) AND  (x1 = TRUE) AND  (x2 = FALSE) AND  (t0.Q = TRUE)) THEN 
        cstate58 := 6338; y0 := FALSE; y1 := FALSE; t0_start := FALSE; 
    ELSIF ((x0 = FALSE) AND  (x1 = TRUE) AND  (x2 = TRUE) AND  (t0.Q = FALSE)) THEN 
        cstate58 := 6532; y0 := FALSE; y1 := FALSE; t0_start := FALSE; 
    ELSIF ((x0 = FALSE) AND  (x1 = TRUE) AND  (x2 = TRUE) AND  (t0.Q = TRUE)) THEN 
        cstate58 := 6530; y0 := FALSE; y1 := FALSE; t0_start := FALSE; 
    ELSIF ((x0 = TRUE) AND  (x1 = FALSE) AND  (x2 = FALSE) AND  (t0.Q = FALSE)) THEN 
        cstate58 := 4168; y0 := TRUE; y1 := FALSE; t0_start := FALSE; 
    ELSIF ((x0 = TRUE) AND  (x1 = FALSE) AND  (x2 = FALSE) AND  (t0.Q = TRUE)) THEN 
        cstate58 := 4162; y0 := TRUE; y1 := FALSE; t0_start := FALSE; 
    ELSIF ((x0 = TRUE) AND  (x1 = FALSE) AND  (x2 = TRUE) AND  (t0.Q = FALSE)) THEN 
        cstate58 := 2824; y0 := FALSE; y1 := FALSE; t0_start := FALSE; 
    ELSIF ((x0 = TRUE) AND  (x1 = FALSE) AND  (x2 = TRUE) AND  (t0.Q = TRUE)) THEN 
        cstate58 := 2818; y0 := FALSE; y1 := FALSE; t0_start := FALSE; 
    ELSIF ((x0 = TRUE) AND  (x1 = TRUE) AND  (x2 = FALSE) AND  (t0.Q = FALSE)) THEN 
        cstate58 := 4678; y0 := TRUE; y1 := FALSE; t0_start := FALSE; 
    ELSIF ((x0 = TRUE) AND  (x1 = TRUE) AND  (x2 = FALSE) AND  (t0.Q = TRUE)) THEN 
        cstate58 := 4674; y0 := TRUE; y1 := FALSE; t0_start := FALSE; 
    ELSIF ((x0 = TRUE) AND  (x1 = TRUE) AND  (x2 = TRUE) AND  (t0.Q = FALSE)) THEN 
        cstate58 := 2502; y0 := FALSE; y1 := FALSE; t0_start := FALSE; 
    ELSIF ((x0 = TRUE) AND  (x1 = TRUE) AND  (x2 = TRUE) AND  (t0.Q = TRUE)) THEN 
        cstate58 := 2498; y0 := FALSE; y1 := FALSE; t0_start := FALSE; 
    END_IF;
6532:
    IF ((x0 = FALSE) AND  (x1 = FALSE) AND  (x2 = FALSE) AND  (t0.Q = FALSE)) THEN 
        cstate58 := 6340; y0 := FALSE; y1 := FALSE; t0_start := FALSE; 
    ELSIF ((x0 = FALSE) AND  (x1 = FALSE) AND  (x2 = FALSE) AND  (t0.Q = TRUE)) THEN 
        cstate58 := 6346; y0 := FALSE; y1 := TRUE; t0_start := FALSE; 
    ELSIF ((x0 = FALSE) AND  (x1 = FALSE) AND  (x2 = TRUE) AND  (t0.Q = FALSE)) THEN 
        cstate58 := 6532; y0 := FALSE; y1 := FALSE; t0_start := FALSE; 
    ELSIF ((x0 = FALSE) AND  (x1 = FALSE) AND  (x2 = TRUE) AND  (t0.Q = TRUE)) THEN 
        cstate58 := 6538; y0 := FALSE; y1 := TRUE; t0_start := FALSE; 
    ELSIF ((x0 = FALSE) AND  (x1 = TRUE) AND  (x2 = FALSE) AND  (t0.Q = FALSE)) THEN 
        cstate58 := 6340; y0 := FALSE; y1 := FALSE; t0_start := FALSE; 
    ELSIF ((x0 = FALSE) AND  (x1 = TRUE) AND  (x2 = FALSE) AND  (t0.Q = TRUE)) THEN 
        cstate58 := 6338; y0 := FALSE; y1 := FALSE; t0_start := FALSE; 
    ELSIF ((x0 = FALSE) AND  (x1 = TRUE) AND  (x2 = TRUE) AND  (t0.Q = FALSE)) THEN 
        cstate58 := 6532; y0 := FALSE; y1 := FALSE; t0_start := FALSE; 
    ELSIF ((x0 = FALSE) AND  (x1 = TRUE) AND  (x2 = TRUE) AND  (t0.Q = TRUE)) THEN 
        cstate58 := 6530; y0 := FALSE; y1 := FALSE; t0_start := FALSE; 
    ELSIF ((x0 = TRUE) AND  (x1 = FALSE) AND  (x2 = FALSE) AND  (t0.Q = FALSE)) THEN 
        cstate58 := 4168; y0 := TRUE; y1 := FALSE; t0_start := FALSE; 
    ELSIF ((x0 = TRUE) AND  (x1 = FALSE) AND  (x2 = FALSE) AND  (t0.Q = TRUE)) THEN 
        cstate58 := 4162; y0 := TRUE; y1 := FALSE; t0_start := FALSE; 
    ELSIF ((x0 = TRUE) AND  (x1 = FALSE) AND  (x2 = TRUE) AND  (t0.Q = FALSE)) THEN 
        cstate58 := 2824; y0 := FALSE; y1 := FALSE; t0_start := FALSE; 
    ELSIF ((x0 = TRUE) AND  (x1 = FALSE) AND  (x2 = TRUE) AND  (t0.Q = TRUE)) THEN 
        cstate58 := 2818; y0 := FALSE; y1 := FALSE; t0_start := FALSE; 
    ELSIF ((x0 = TRUE) AND  (x1 = TRUE) AND  (x2 = FALSE) AND  (t0.Q = FALSE)) THEN 
        cstate58 := 4678; y0 := TRUE; y1 := FALSE; t0_start := FALSE; 
    ELSIF ((x0 = TRUE) AND  (x1 = TRUE) AND  (x2 = FALSE) AND  (t0.Q = TRUE)) THEN 
        cstate58 := 4674; y0 := TRUE; y1 := FALSE; t0_start := FALSE; 
    ELSIF ((x0 = TRUE) AND  (x1 = TRUE) AND  (x2 = TRUE) AND  (t0.Q = FALSE)) THEN 
        cstate58 := 2502; y0 := FALSE; y1 := FALSE; t0_start := FALSE; 
    ELSIF ((x0 = TRUE) AND  (x1 = TRUE) AND  (x2 = TRUE) AND  (t0.Q = TRUE)) THEN 
        cstate58 := 2498; y0 := FALSE; y1 := FALSE; t0_start := FALSE; 
    END_IF;
7364:
    IF ((x0 = FALSE) AND  (x1 = FALSE) AND  (x2 = FALSE) AND  (t0.Q = FALSE)) THEN 
        cstate58 := 7364; y0 := FALSE; y1 := FALSE; t0_start := FALSE; 
    ELSIF ((x0 = FALSE) AND  (x1 = FALSE) AND  (x2 = FALSE) AND  (t0.Q = TRUE)) THEN 
        cstate58 := 7370; y0 := FALSE; y1 := TRUE; t0_start := FALSE; 
    ELSIF ((x0 = FALSE) AND  (x1 = FALSE) AND  (x2 = TRUE) AND  (t0.Q = FALSE)) THEN 
        cstate58 := 7492; y0 := FALSE; y1 := FALSE; t0_start := TRUE; t0_up := FALSE; 
    ELSIF ((x0 = FALSE) AND  (x1 = FALSE) AND  (x2 = TRUE) AND  (t0.Q = TRUE)) THEN 
        cstate58 := 7500; y0 := FALSE; y1 := TRUE; t0_start := TRUE; t0_up := FALSE; 
    ELSIF ((x0 = FALSE) AND  (x1 = TRUE) AND  (x2 = FALSE) AND  (t0.Q = FALSE)) THEN 
        cstate58 := 6340; y0 := FALSE; y1 := FALSE; t0_start := FALSE; 
    ELSIF ((x0 = FALSE) AND  (x1 = TRUE) AND  (x2 = FALSE) AND  (t0.Q = TRUE)) THEN 
        cstate58 := 6338; y0 := FALSE; y1 := FALSE; t0_start := FALSE; 
    ELSIF ((x0 = FALSE) AND  (x1 = TRUE) AND  (x2 = TRUE) AND  (t0.Q = FALSE)) THEN 
        cstate58 := 6468; y0 := FALSE; y1 := FALSE; t0_start := TRUE; t0_up := FALSE; 
    ELSIF ((x0 = FALSE) AND  (x1 = TRUE) AND  (x2 = TRUE) AND  (t0.Q = TRUE)) THEN 
        cstate58 := 6466; y0 := FALSE; y1 := FALSE; t0_start := TRUE; t0_up := FALSE; 
    ELSIF ((x0 = TRUE) AND  (x1 = FALSE) AND  (x2 = FALSE) AND  (t0.Q = FALSE)) THEN 
        cstate58 := 5192; y0 := TRUE; y1 := FALSE; t0_start := FALSE; 
    ELSIF ((x0 = TRUE) AND  (x1 = FALSE) AND  (x2 = FALSE) AND  (t0.Q = TRUE)) THEN 
        cstate58 := 5186; y0 := TRUE; y1 := FALSE; t0_start := FALSE; 
    ELSIF ((x0 = TRUE) AND  (x1 = FALSE) AND  (x2 = TRUE) AND  (t0.Q = FALSE)) THEN 
        cstate58 := 3784; y0 := FALSE; y1 := FALSE; t0_start := TRUE; t0_up := FALSE; 
    ELSIF ((x0 = TRUE) AND  (x1 = FALSE) AND  (x2 = TRUE) AND  (t0.Q = TRUE)) THEN 
        cstate58 := 3778; y0 := FALSE; y1 := FALSE; t0_start := TRUE; t0_up := FALSE; 
    ELSIF ((x0 = TRUE) AND  (x1 = TRUE) AND  (x2 = FALSE) AND  (t0.Q = FALSE)) THEN 
        cstate58 := 4678; y0 := TRUE; y1 := FALSE; t0_start := FALSE; 
    ELSIF ((x0 = TRUE) AND  (x1 = TRUE) AND  (x2 = FALSE) AND  (t0.Q = TRUE)) THEN 
        cstate58 := 4674; y0 := TRUE; y1 := FALSE; t0_start := FALSE; 
    ELSIF ((x0 = TRUE) AND  (x1 = TRUE) AND  (x2 = TRUE) AND  (t0.Q = FALSE)) THEN 
        cstate58 := 2566; y0 := FALSE; y1 := FALSE; t0_start := TRUE; t0_up := FALSE; 
    ELSIF ((x0 = TRUE) AND  (x1 = TRUE) AND  (x2 = TRUE) AND  (t0.Q = TRUE)) THEN 
        cstate58 := 2562; y0 := FALSE; y1 := FALSE; t0_start := TRUE; t0_up := FALSE; 
    END_IF;
6428:
    IF ((x0 = FALSE) AND  (x1 = FALSE) AND  (x2 = FALSE) AND  (t0.Q = FALSE)) THEN 
        cstate58 := 6428; y0 := FALSE; y1 := TRUE; t0_start := FALSE; 
    ELSIF ((x0 = FALSE) AND  (x1 = FALSE) AND  (x2 = FALSE) AND  (t0.Q = TRUE)) THEN 
        cstate58 := 6350; y0 := FALSE; y1 := TRUE; t0_start := FALSE; 
    ELSIF ((x0 = FALSE) AND  (x1 = FALSE) AND  (x2 = TRUE) AND  (t0.Q = FALSE)) THEN 
        cstate58 := 6492; y0 := FALSE; y1 := TRUE; t0_start := TRUE; t0_up := FALSE; 
    ELSIF ((x0 = FALSE) AND  (x1 = FALSE) AND  (x2 = TRUE) AND  (t0.Q = TRUE)) THEN 
        cstate58 := 6480; y0 := FALSE; y1 := TRUE; t0_start := TRUE; t0_up := FALSE; 
    ELSIF ((x0 = FALSE) AND  (x1 = TRUE) AND  (x2 = FALSE) AND  (t0.Q = FALSE)) THEN 
        cstate58 := 6404; y0 := FALSE; y1 := FALSE; t0_start := FALSE; 
    ELSIF ((x0 = FALSE) AND  (x1 = TRUE) AND  (x2 = FALSE) AND  (t0.Q = TRUE)) THEN 
        cstate58 := 6338; y0 := FALSE; y1 := FALSE; t0_start := FALSE; 
    ELSIF ((x0 = FALSE) AND  (x1 = TRUE) AND  (x2 = TRUE) AND  (t0.Q = FALSE)) THEN 
        cstate58 := 6468; y0 := FALSE; y1 := FALSE; t0_start := TRUE; t0_up := FALSE; 
    ELSIF ((x0 = FALSE) AND  (x1 = TRUE) AND  (x2 = TRUE) AND  (t0.Q = TRUE)) THEN 
        cstate58 := 6466; y0 := FALSE; y1 := FALSE; t0_start := TRUE; t0_up := FALSE; 
    ELSIF ((x0 = TRUE) AND  (x1 = FALSE) AND  (x2 = FALSE) AND  (t0.Q = FALSE)) THEN 
        cstate58 := 4232; y0 := TRUE; y1 := FALSE; t0_start := FALSE; 
    ELSIF ((x0 = TRUE) AND  (x1 = FALSE) AND  (x2 = FALSE) AND  (t0.Q = TRUE)) THEN 
        cstate58 := 4162; y0 := TRUE; y1 := FALSE; t0_start := FALSE; 
    ELSIF ((x0 = TRUE) AND  (x1 = FALSE) AND  (x2 = TRUE) AND  (t0.Q = FALSE)) THEN 
        cstate58 := 2760; y0 := FALSE; y1 := FALSE; t0_start := TRUE; t0_up := FALSE; 
    ELSIF ((x0 = TRUE) AND  (x1 = FALSE) AND  (x2 = TRUE) AND  (t0.Q = TRUE)) THEN 
        cstate58 := 2754; y0 := FALSE; y1 := FALSE; t0_start := TRUE; t0_up := FALSE; 
    ELSIF ((x0 = TRUE) AND  (x1 = TRUE) AND  (x2 = FALSE) AND  (t0.Q = FALSE)) THEN 
        cstate58 := 4742; y0 := TRUE; y1 := FALSE; t0_start := FALSE; 
    ELSIF ((x0 = TRUE) AND  (x1 = TRUE) AND  (x2 = FALSE) AND  (t0.Q = TRUE)) THEN 
        cstate58 := 4674; y0 := TRUE; y1 := FALSE; t0_start := FALSE; 
    ELSIF ((x0 = TRUE) AND  (x1 = TRUE) AND  (x2 = TRUE) AND  (t0.Q = FALSE)) THEN 
        cstate58 := 2566; y0 := FALSE; y1 := FALSE; t0_start := TRUE; t0_up := FALSE; 
    ELSIF ((x0 = TRUE) AND  (x1 = TRUE) AND  (x2 = TRUE) AND  (t0.Q = TRUE)) THEN 
        cstate58 := 2562; y0 := FALSE; y1 := FALSE; t0_start := TRUE; t0_up := FALSE; 
    END_IF;
7362:
    IF ((x0 = FALSE) AND  (x1 = FALSE) AND  (x2 = FALSE) AND  (t0.Q = FALSE)) THEN 
        cstate58 := 7364; y0 := FALSE; y1 := FALSE; t0_start := FALSE; 
    ELSIF ((x0 = FALSE) AND  (x1 = FALSE) AND  (x2 = FALSE) AND  (t0.Q = TRUE)) THEN 
        cstate58 := 7362; y0 := FALSE; y1 := FALSE; t0_start := FALSE; 
    ELSIF ((x0 = FALSE) AND  (x1 = FALSE) AND  (x2 = TRUE) AND  (t0.Q = FALSE)) THEN 
        cstate58 := 7492; y0 := FALSE; y1 := FALSE; t0_start := TRUE; t0_up := FALSE; 
    ELSIF ((x0 = FALSE) AND  (x1 = FALSE) AND  (x2 = TRUE) AND  (t0.Q = TRUE)) THEN 
        cstate58 := 7490; y0 := FALSE; y1 := FALSE; t0_start := TRUE; t0_up := FALSE; 
    ELSIF ((x0 = FALSE) AND  (x1 = TRUE) AND  (x2 = FALSE) AND  (t0.Q = FALSE)) THEN 
        cstate58 := 6340; y0 := FALSE; y1 := FALSE; t0_start := FALSE; 
    ELSIF ((x0 = FALSE) AND  (x1 = TRUE) AND  (x2 = FALSE) AND  (t0.Q = TRUE)) THEN 
        cstate58 := 6338; y0 := FALSE; y1 := FALSE; t0_start := FALSE; 
    ELSIF ((x0 = FALSE) AND  (x1 = TRUE) AND  (x2 = TRUE) AND  (t0.Q = FALSE)) THEN 
        cstate58 := 6468; y0 := FALSE; y1 := FALSE; t0_start := TRUE; t0_up := FALSE; 
    ELSIF ((x0 = FALSE) AND  (x1 = TRUE) AND  (x2 = TRUE) AND  (t0.Q = TRUE)) THEN 
        cstate58 := 6466; y0 := FALSE; y1 := FALSE; t0_start := TRUE; t0_up := FALSE; 
    ELSIF ((x0 = TRUE) AND  (x1 = FALSE) AND  (x2 = FALSE) AND  (t0.Q = FALSE)) THEN 
        cstate58 := 5192; y0 := TRUE; y1 := FALSE; t0_start := FALSE; 
    ELSIF ((x0 = TRUE) AND  (x1 = FALSE) AND  (x2 = FALSE) AND  (t0.Q = TRUE)) THEN 
        cstate58 := 5186; y0 := TRUE; y1 := FALSE; t0_start := FALSE; 
    ELSIF ((x0 = TRUE) AND  (x1 = FALSE) AND  (x2 = TRUE) AND  (t0.Q = FALSE)) THEN 
        cstate58 := 3784; y0 := FALSE; y1 := FALSE; t0_start := TRUE; t0_up := FALSE; 
    ELSIF ((x0 = TRUE) AND  (x1 = FALSE) AND  (x2 = TRUE) AND  (t0.Q = TRUE)) THEN 
        cstate58 := 3778; y0 := FALSE; y1 := FALSE; t0_start := TRUE; t0_up := FALSE; 
    ELSIF ((x0 = TRUE) AND  (x1 = TRUE) AND  (x2 = FALSE) AND  (t0.Q = FALSE)) THEN 
        cstate58 := 4678; y0 := TRUE; y1 := FALSE; t0_start := FALSE; 
    ELSIF ((x0 = TRUE) AND  (x1 = TRUE) AND  (x2 = FALSE) AND  (t0.Q = TRUE)) THEN 
        cstate58 := 4674; y0 := TRUE; y1 := FALSE; t0_start := FALSE; 
    ELSIF ((x0 = TRUE) AND  (x1 = TRUE) AND  (x2 = TRUE) AND  (t0.Q = FALSE)) THEN 
        cstate58 := 2566; y0 := FALSE; y1 := FALSE; t0_start := TRUE; t0_up := FALSE; 
    ELSIF ((x0 = TRUE) AND  (x1 = TRUE) AND  (x2 = TRUE) AND  (t0.Q = TRUE)) THEN 
        cstate58 := 2562; y0 := FALSE; y1 := FALSE; t0_start := TRUE; t0_up := FALSE; 
    END_IF;
1356:
    IF ((x0 = FALSE) AND  (x1 = FALSE) AND  (x2 = FALSE) AND  (t0.Q = FALSE)) THEN 
        cstate58 := 1304; y0 := FALSE; y1 := TRUE; t0_start := FALSE; 
    ELSIF ((x0 = FALSE) AND  (x1 = FALSE) AND  (x2 = FALSE) AND  (t0.Q = TRUE)) THEN 
        cstate58 := 1226; y0 := FALSE; y1 := TRUE; t0_start := FALSE; 
    ELSIF ((x0 = FALSE) AND  (x1 = FALSE) AND  (x2 = TRUE) AND  (t0.Q = FALSE)) THEN 
        cstate58 := 1368; y0 := FALSE; y1 := TRUE; t0_start := FALSE; 
    ELSIF ((x0 = FALSE) AND  (x1 = FALSE) AND  (x2 = TRUE) AND  (t0.Q = TRUE)) THEN 
        cstate58 := 1418; y0 := FALSE; y1 := TRUE; t0_start := FALSE; 
    ELSIF ((x0 = FALSE) AND  (x1 = TRUE) AND  (x2 = FALSE) AND  (t0.Q = FALSE)) THEN 
        cstate58 := 1284; y0 := FALSE; y1 := FALSE; t0_start := FALSE; 
    ELSIF ((x0 = FALSE) AND  (x1 = TRUE) AND  (x2 = FALSE) AND  (t0.Q = TRUE)) THEN 
        cstate58 := 1218; y0 := FALSE; y1 := FALSE; t0_start := FALSE; 
    ELSIF ((x0 = FALSE) AND  (x1 = TRUE) AND  (x2 = TRUE) AND  (t0.Q = FALSE)) THEN 
        cstate58 := 1348; y0 := FALSE; y1 := FALSE; t0_start := FALSE; 
    ELSIF ((x0 = FALSE) AND  (x1 = TRUE) AND  (x2 = TRUE) AND  (t0.Q = TRUE)) THEN 
        cstate58 := 1410; y0 := FALSE; y1 := FALSE; t0_start := FALSE; 
    ELSIF ((x0 = TRUE) AND  (x1 = FALSE) AND  (x2 = FALSE) AND  (t0.Q = FALSE)) THEN 
        cstate58 := 5256; y0 := TRUE; y1 := FALSE; t0_start := FALSE; 
    ELSIF ((x0 = TRUE) AND  (x1 = FALSE) AND  (x2 = FALSE) AND  (t0.Q = TRUE)) THEN 
        cstate58 := 5186; y0 := TRUE; y1 := FALSE; t0_start := FALSE; 
    ELSIF ((x0 = TRUE) AND  (x1 = FALSE) AND  (x2 = TRUE) AND  (t0.Q = FALSE)) THEN 
        cstate58 := 3784; y0 := FALSE; y1 := FALSE; t0_start := FALSE; 
    ELSIF ((x0 = TRUE) AND  (x1 = FALSE) AND  (x2 = TRUE) AND  (t0.Q = TRUE)) THEN 
        cstate58 := 3842; y0 := FALSE; y1 := FALSE; t0_start := FALSE; 
    ELSIF ((x0 = TRUE) AND  (x1 = TRUE) AND  (x2 = FALSE) AND  (t0.Q = FALSE)) THEN 
        cstate58 := 4742; y0 := TRUE; y1 := FALSE; t0_start := FALSE; 
    ELSIF ((x0 = TRUE) AND  (x1 = TRUE) AND  (x2 = FALSE) AND  (t0.Q = TRUE)) THEN 
        cstate58 := 4674; y0 := TRUE; y1 := FALSE; t0_start := FALSE; 
    ELSIF ((x0 = TRUE) AND  (x1 = TRUE) AND  (x2 = TRUE) AND  (t0.Q = FALSE)) THEN 
        cstate58 := 2566; y0 := FALSE; y1 := FALSE; t0_start := FALSE; 
    ELSIF ((x0 = TRUE) AND  (x1 = TRUE) AND  (x2 = TRUE) AND  (t0.Q = TRUE)) THEN 
        cstate58 := 2498; y0 := FALSE; y1 := FALSE; t0_start := FALSE; 
    END_IF;
1218:
    IF ((x0 = FALSE) AND  (x1 = FALSE) AND  (x2 = FALSE) AND  (t0.Q = FALSE)) THEN 
        cstate58 := 1220; y0 := FALSE; y1 := FALSE; t0_start := FALSE; 
    ELSIF ((x0 = FALSE) AND  (x1 = FALSE) AND  (x2 = FALSE) AND  (t0.Q = TRUE)) THEN 
        cstate58 := 1218; y0 := FALSE; y1 := FALSE; t0_start := FALSE; 
    ELSIF ((x0 = FALSE) AND  (x1 = FALSE) AND  (x2 = TRUE) AND  (t0.Q = FALSE)) THEN 
        cstate58 := 1348; y0 := FALSE; y1 := FALSE; t0_start := TRUE; t0_up := FALSE; 
    ELSIF ((x0 = FALSE) AND  (x1 = FALSE) AND  (x2 = TRUE) AND  (t0.Q = TRUE)) THEN 
        cstate58 := 1346; y0 := FALSE; y1 := FALSE; t0_start := TRUE; t0_up := FALSE; 
    ELSIF ((x0 = FALSE) AND  (x1 = TRUE) AND  (x2 = FALSE) AND  (t0.Q = FALSE)) THEN 
        cstate58 := 1220; y0 := FALSE; y1 := FALSE; t0_start := FALSE; 
    ELSIF ((x0 = FALSE) AND  (x1 = TRUE) AND  (x2 = FALSE) AND  (t0.Q = TRUE)) THEN 
        cstate58 := 1218; y0 := FALSE; y1 := FALSE; t0_start := FALSE; 
    ELSIF ((x0 = FALSE) AND  (x1 = TRUE) AND  (x2 = TRUE) AND  (t0.Q = FALSE)) THEN 
        cstate58 := 1348; y0 := FALSE; y1 := FALSE; t0_start := TRUE; t0_up := FALSE; 
    ELSIF ((x0 = FALSE) AND  (x1 = TRUE) AND  (x2 = TRUE) AND  (t0.Q = TRUE)) THEN 
        cstate58 := 1346; y0 := FALSE; y1 := FALSE; t0_start := TRUE; t0_up := FALSE; 
    ELSIF ((x0 = TRUE) AND  (x1 = FALSE) AND  (x2 = FALSE) AND  (t0.Q = FALSE)) THEN 
        cstate58 := 5192; y0 := TRUE; y1 := FALSE; t0_start := FALSE; 
    ELSIF ((x0 = TRUE) AND  (x1 = FALSE) AND  (x2 = FALSE) AND  (t0.Q = TRUE)) THEN 
        cstate58 := 5186; y0 := TRUE; y1 := FALSE; t0_start := FALSE; 
    ELSIF ((x0 = TRUE) AND  (x1 = FALSE) AND  (x2 = TRUE) AND  (t0.Q = FALSE)) THEN 
        cstate58 := 3784; y0 := FALSE; y1 := FALSE; t0_start := TRUE; t0_up := FALSE; 
    ELSIF ((x0 = TRUE) AND  (x1 = FALSE) AND  (x2 = TRUE) AND  (t0.Q = TRUE)) THEN 
        cstate58 := 3778; y0 := FALSE; y1 := FALSE; t0_start := TRUE; t0_up := FALSE; 
    ELSIF ((x0 = TRUE) AND  (x1 = TRUE) AND  (x2 = FALSE) AND  (t0.Q = FALSE)) THEN 
        cstate58 := 4678; y0 := TRUE; y1 := FALSE; t0_start := FALSE; 
    ELSIF ((x0 = TRUE) AND  (x1 = TRUE) AND  (x2 = FALSE) AND  (t0.Q = TRUE)) THEN 
        cstate58 := 4674; y0 := TRUE; y1 := FALSE; t0_start := FALSE; 
    ELSIF ((x0 = TRUE) AND  (x1 = TRUE) AND  (x2 = TRUE) AND  (t0.Q = FALSE)) THEN 
        cstate58 := 2566; y0 := FALSE; y1 := FALSE; t0_start := TRUE; t0_up := FALSE; 
    ELSIF ((x0 = TRUE) AND  (x1 = TRUE) AND  (x2 = TRUE) AND  (t0.Q = TRUE)) THEN 
        cstate58 := 2562; y0 := FALSE; y1 := FALSE; t0_start := TRUE; t0_up := FALSE; 
    END_IF;
6424:
    IF ((x0 = FALSE) AND  (x1 = FALSE) AND  (x2 = FALSE) AND  (t0.Q = FALSE)) THEN 
        cstate58 := 6424; y0 := FALSE; y1 := TRUE; t0_start := FALSE; 
    ELSIF ((x0 = FALSE) AND  (x1 = FALSE) AND  (x2 = FALSE) AND  (t0.Q = TRUE)) THEN 
        cstate58 := 6346; y0 := FALSE; y1 := TRUE; t0_start := FALSE; 
    ELSIF ((x0 = FALSE) AND  (x1 = FALSE) AND  (x2 = TRUE) AND  (t0.Q = FALSE)) THEN 
        cstate58 := 6488; y0 := FALSE; y1 := TRUE; t0_start := TRUE; t0_up := FALSE; 
    ELSIF ((x0 = FALSE) AND  (x1 = FALSE) AND  (x2 = TRUE) AND  (t0.Q = TRUE)) THEN 
        cstate58 := 6476; y0 := FALSE; y1 := TRUE; t0_start := TRUE; t0_up := FALSE; 
    ELSIF ((x0 = FALSE) AND  (x1 = TRUE) AND  (x2 = FALSE) AND  (t0.Q = FALSE)) THEN 
        cstate58 := 6404; y0 := FALSE; y1 := FALSE; t0_start := FALSE; 
    ELSIF ((x0 = FALSE) AND  (x1 = TRUE) AND  (x2 = FALSE) AND  (t0.Q = TRUE)) THEN 
        cstate58 := 6338; y0 := FALSE; y1 := FALSE; t0_start := FALSE; 
    ELSIF ((x0 = FALSE) AND  (x1 = TRUE) AND  (x2 = TRUE) AND  (t0.Q = FALSE)) THEN 
        cstate58 := 6468; y0 := FALSE; y1 := FALSE; t0_start := TRUE; t0_up := FALSE; 
    ELSIF ((x0 = FALSE) AND  (x1 = TRUE) AND  (x2 = TRUE) AND  (t0.Q = TRUE)) THEN 
        cstate58 := 6466; y0 := FALSE; y1 := FALSE; t0_start := TRUE; t0_up := FALSE; 
    ELSIF ((x0 = TRUE) AND  (x1 = FALSE) AND  (x2 = FALSE) AND  (t0.Q = FALSE)) THEN 
        cstate58 := 4232; y0 := TRUE; y1 := FALSE; t0_start := FALSE; 
    ELSIF ((x0 = TRUE) AND  (x1 = FALSE) AND  (x2 = FALSE) AND  (t0.Q = TRUE)) THEN 
        cstate58 := 4162; y0 := TRUE; y1 := FALSE; t0_start := FALSE; 
    ELSIF ((x0 = TRUE) AND  (x1 = FALSE) AND  (x2 = TRUE) AND  (t0.Q = FALSE)) THEN 
        cstate58 := 2760; y0 := FALSE; y1 := FALSE; t0_start := TRUE; t0_up := FALSE; 
    ELSIF ((x0 = TRUE) AND  (x1 = FALSE) AND  (x2 = TRUE) AND  (t0.Q = TRUE)) THEN 
        cstate58 := 2754; y0 := FALSE; y1 := FALSE; t0_start := TRUE; t0_up := FALSE; 
    ELSIF ((x0 = TRUE) AND  (x1 = TRUE) AND  (x2 = FALSE) AND  (t0.Q = FALSE)) THEN 
        cstate58 := 4742; y0 := TRUE; y1 := FALSE; t0_start := FALSE; 
    ELSIF ((x0 = TRUE) AND  (x1 = TRUE) AND  (x2 = FALSE) AND  (t0.Q = TRUE)) THEN 
        cstate58 := 4674; y0 := TRUE; y1 := FALSE; t0_start := FALSE; 
    ELSIF ((x0 = TRUE) AND  (x1 = TRUE) AND  (x2 = TRUE) AND  (t0.Q = FALSE)) THEN 
        cstate58 := 2566; y0 := FALSE; y1 := FALSE; t0_start := TRUE; t0_up := FALSE; 
    ELSIF ((x0 = TRUE) AND  (x1 = TRUE) AND  (x2 = TRUE) AND  (t0.Q = TRUE)) THEN 
        cstate58 := 2562; y0 := FALSE; y1 := FALSE; t0_start := TRUE; t0_up := FALSE; 
    END_IF;
END_CASE;

(* Additional processing to handle clocks - in CODESYS, it only starts
    with rising edge and can not be placed inside IF statement *) 
IF(t0_up = TRUE) THEN
    t0_reset := TRUE;
ELSIF(t0_start = TRUE AND t0_up = FALSE) THEN
    t0_up := TRUE;  t0_reset := FALSE;
END_IF
t0(IN:=t0_reset, PT:=T0_VALUE);

END_FUNCTION_BLOCK
